(* IEC 61131-3 sources: trust-platform/crates/trust-runtime/tests/fixtures/plcopen_motion/single_axis_negative_transition_vel_next/src, 1 file *)

(* ---- tests.st ---- *)
PROGRAM plcopen_motion_single_axis_negative_transition_vel_next
VAR
    WrongBufferMode : MC_BUFFER_MODE;
END_VAR

WrongBufferMode := MC_BUFFER_MODE#mcTransitionVelNext;
END_PROGRAM
